Fanuc KAREL source: kc00019.KL

-- PROVISIONAL review KL for V940-1; original PC SHA256 a2daed3f837e3e17818bc099d00c12571706b262eea0a9a175f9ecded389d1e9
-- Incomplete behavior may be omitted. Consult companion uncertainty JSON. Do not deploy.
PROGRAM KC00019
%NOLOCKGROUP
BEGIN
  -- V9_ZERO_TABLE_METADATA_HINT layout=0002_ascii; no indexed target words; source/name/runtime held
  -- UNRESOLVED_PC offsets 5-53; opcodes 27,22,22,22,22,22,2A,22,22,31
  -- UNRESOLVED_PC offsets 58-62; opcodes 7F
END KC00019
